(* IEC 61131-3 sources: Lasal-MCP/examples/SampleSource/4_PumpControlSchemeSolution/Stations/MachineControl/MachineControl/Class/PumpControl, 1 file *)

(* ---- PumpControl.st ---- *)
(*!
<Class
	Name               = "PumpControl"
	Revision           = "0.0"
	RealtimeTask       = "false"
	CyclicTask         = "true"
	DefCyclictime      = "10 ms"
	BackgroundTask     = "false"
	Sigmatek           = "false"
	OSInterface        = "false"
	HighPriority       = "false"
	Automatic          = "false"
	UpdateMode         = "Prescan"
	SharedCommandTable = "true"
	Objectsize         = "(630,540)">
	<Channels>
		<Server Name="ActFillLevelVisu" Visualized="true" Initialize="false" WriteProtected="true" Retentive="false"/>
		<Server Name="MaxAlarm" Visualized="true" Initialize="true" DefValue="45000" WriteProtected="false" Retentive="File"/>
		<Server Name="MaxBorder" Visualized="true" Initialize="true" DefValue="40000" WriteProtected="false" Retentive="File"/>
		<Server Name="MinAlarm" Visualized="true" Initialize="true" DefValue="5000" WriteProtected="false" Retentive="File"/>
		<Server Name="MinBorder" Visualized="true" Initialize="true" DefValue="10000" WriteProtected="false" Retentive="File"/>
		<Server Name="PumpControlName" Visualized="true" Remotely="true" Initialize="true" WriteProtected="false" Retentive="File"/>
		<Server Name="PumpVisu" Visualized="true" Initialize="false" WriteProtected="true" Retentive="false"/>
		<Server Name="WaterTempVisu" Visualized="true" Initialize="false" WriteProtected="true" Retentive="false"/>
		<Client Name="_AlarmX1Para1" Required="true" Internal="true"/>
		<Client Name="_AlarmX1Para2" Required="true" Internal="true"/>
		<Client Name="_AlarmX2Para1" Required="true" Internal="true"/>
		<Client Name="ActFillLevel" Required="true" Internal="false"/>
		<Client Name="Pump" Required="true" Internal="false"/>
		<Client Name="StringRAM1" Required="true" Internal="true"/>
		<Client Name="WaterTemp" Required="true" Internal="false"/>
	</Channels>
	<Network Name="PumpControl">
		<!-- List of Components in this network -->
		<Components>
			<Object
				Name       = "_AlarmX1Para1"
				Class      = "_AlarmX1Para"
				Position   = "(470,570)"
				Visualized = "true"
				Remotely   = "true">
				<Channels>
					<Server Name="ClassSvr"/>
					<Client Name="Acknow"/>
					<Client Name="Config" Value="0"/>
					<Client Name="Group"/>
					<Client Name="Para1"/>
				</Channels>
			</Object>
			<Object
				Name       = "_AlarmX1Para2"
				Class      = "_AlarmX1Para"
				Position   = "(470,900)"
				Visualized = "true"
				Remotely   = "true">
				<Channels>
					<Server Name="ClassSvr"/>
					<Client Name="Acknow"/>
					<Client Name="Config" Value="0"/>
					<Client Name="Group"/>
					<Client Name="Para1"/>
				</Channels>
			</Object>
			<Object
				Name       = "_AlarmX2Para1"
				Class      = "_AlarmX2Para"
				Position   = "(470,1230)"
				Visualized = "true"
				Remotely   = "true">
				<Channels>
					<Server Name="ClassSvr"/>
					<Client Name="Acknow"/>
					<Client Name="Config" Value="0"/>
					<Client Name="Group"/>
					<Client Name="Para1" Value="0"/>
					<Client Name="Para2"/>
				</Channels>
			</Object>
			<Object
				Name       = "StringRAM1"
				Class      = "StringRAM"
				Position   = "(470,1620)"
				Visualized = "true"
				Remotely   = "true">
				<Channels>
					<Server Name="Data"/>
					<Client Name="SingleRealloc" Value="1"/>
					<Client Name="UseFile"/>
				</Channels>
			</Object>
		</Components>
		<Comments>
		</Comments>
		<!-- List of Connections in this network -->
		<Connections>
			<Connection Source="this._AlarmX1Para1" Destination="_AlarmX1Para1.ClassSvr"/>
			<Connection Source="this._AlarmX1Para2" Destination="_AlarmX1Para2.ClassSvr"/>
			<Connection Source="this._AlarmX2Para1" Destination="_AlarmX2Para1.ClassSvr"/>
			<Connection Source="this.StringRAM1" Destination="StringRAM1.Data"/>
			<Connection Source="this.PumpControlName" Destination="StringRAM1.Data" Vertices="(1048,630),(876,1710),"/>
		</Connections>
		<!-- Headerfiles -->
		<Options>
		</Options>
	</Network>
</Class>
*)
PumpControl : CLASS
  //Servers:
	MaxBorder 	: SvrChCmd_DINT;
	MinBorder 	: SvrCh_DINT;
	MaxAlarm 	: SvrCh_DINT;
	MinAlarm 	: SvrCh_DINT;
	ActFillLevelVisu 	: SvrCh_DINT;
	PumpVisu 	: SvrCh_DINT;
	WaterTempVisu 	: SvrCh_DINT;
	PumpControlName 	: SvrCh_UDINT;
  //Clients:
	ActFillLevel 	: CltCh_DINT;
	Pump 	: CltCh_DINT;
	_AlarmX1Para1 	: CltChCmd__AlarmX1Para;
	_AlarmX1Para2 	: CltChCmd__AlarmX1Para;
	_AlarmX2Para1 	: CltChCmd__AlarmX2Para;
	WaterTemp 	: CltCh_DINT;
	StringRAM1 	: CltChCmd_StringRAM;
  //Variables:
  //Functions:

	FUNCTION VIRTUAL GLOBAL CyWork
		VAR_INPUT
			EAX 	: UDINT;
		END_VAR
		VAR_OUTPUT
			state (EAX) 	: UDINT;
		END_VAR;

	FUNCTION VIRTUAL GLOBAL ActFillLevelVisu::Read
		VAR_OUTPUT
			output (EAX) 	: DINT;
		END_VAR;

	FUNCTION VIRTUAL GLOBAL PumpVisu::Read
		VAR_OUTPUT
			output (EAX) 	: DINT;
		END_VAR;

	FUNCTION VIRTUAL GLOBAL WaterTempVisu::Read
		VAR_OUTPUT
			output (EAX) 	: DINT;
		END_VAR;

	FUNCTION VIRTUAL GLOBAL PumpControlName::Read
		VAR_OUTPUT
			output (EAX) 	: UDINT;
		END_VAR;

	FUNCTION VIRTUAL GLOBAL PumpControlName::Write
		VAR_INPUT
			input (EAX) 	: UDINT;
		END_VAR
		VAR_OUTPUT
			result (EAX) 	: UDINT;
		END_VAR;
  //Tables:
	FUNCTION @STD
		VAR_OUTPUT
			ret_code	: CONFSTATES;
		END_VAR;
	FUNCTION GLOBAL TAB @CT_;
END_CLASS;

#pragma using _AlarmX1Para
#pragma using _AlarmX2Para
#pragma using StringRAM

FUNCTION VIRTUAL GLOBAL PumpControl::CyWork
	VAR_INPUT
		EAX 	: UDINT;
	END_VAR
	VAR_OUTPUT
		state (EAX) 	: UDINT;
	END_VAR

  // read Inputs
  ActFillLevel := ActFillLevel.Read();
  WaterTemp := WaterTemp.Read();

  // Switch off cablebreak
  if ActFillLevel < 0 then
    ActFillLevel := 50000;
  end_if;

  // Alarm Handling
  if ActFillLevel > MaxAlarm then
    _AlarmX1Para1.ClassSvr.Write(input:= 1);
  elsif ActFillLevel < MinAlarm then
    _AlarmX1Para2.ClassSvr.Write(input:= 1);
  else
    _AlarmX1Para1.ClassSvr.Write(input:= 0);
    _AlarmX1Para2.ClassSvr.Write(input:= 0);
  end_if;

  if MaxBorder <= MinBorder then
    _AlarmX2Para1.ClassSvr.Write(input:= 1);
  else
    _AlarmX2Para1.ClassSvr.Write(input:= 0);
  end_if;

  // PumpControl Logic
  if ActFillLevel >= MaxBorder then
    Pump := 1;
  elsif ActFillLevel <= MinBorder then
    Pump := 0;
  end_if;

  // write Outputs
  Pump.Write (Pump);

	state := READY;

END_FUNCTION

FUNCTION VIRTUAL GLOBAL PumpControl::ActFillLevelVisu::Read
	VAR_OUTPUT
		output (EAX) 	: DINT;
	END_VAR

	ActFillLevelVisu := ActFillLevel;

	output := ActFillLevelVisu;

END_FUNCTION

FUNCTION VIRTUAL GLOBAL PumpControl::PumpVisu::Read
	VAR_OUTPUT
		output (EAX) 	: DINT;
	END_VAR

	PumpVisu := Pump;

	output := PumpVisu;

END_FUNCTION

FUNCTION VIRTUAL GLOBAL PumpControl::WaterTempVisu::Read
	VAR_OUTPUT
		output (EAX) 	: DINT;
	END_VAR

	WaterTempVisu := WaterTemp;

	output := WaterTempVisu;

END_FUNCTION

FUNCTION VIRTUAL GLOBAL PumpControl::PumpControlName::Read
	VAR_OUTPUT
		output (EAX) 	: UDINT;
	END_VAR

	PumpControlName := StringRAM1.Data.Read();
	output := PumpControlName;

END_FUNCTION

FUNCTION VIRTUAL GLOBAL PumpControl::PumpControlName::Write
	VAR_INPUT
		input (EAX) 	: UDINT;
	END_VAR
	VAR_OUTPUT
		result (EAX) 	: UDINT;
	END_VAR

	PumpControlName := input;
	result := (StringRAM1.Data.Write(PumpControlName))$UDINT;

END_FUNCTION
